{attribute 'qualified_only'}
VAR_GLOBAL	


END_VAR

(* stored: Version 1.1.0.1
   GVL GVL: Id {b3c39c5b-9457-4b3f-896c-732254fc9b9c} *)
